{attribute 'Tc2GvlVarNames'}
VAR_GLOBAL
	stgGr05HMI			:ST_Gr05HMIRef;
END_VAR

(* stored: Version 1.1.0.1, ProductVersion 3.1.4024.15
   GVL GVL_Gr05HMI: Id {f911afe8-f41c-42c9-827b-d3331d274681} *)
